Staubli VAL3: getTrajList.pgx

public program getTrajList(string& x_sItem[], num x_nIndex)
  local trsf l_tTrsf
  local string l_sItem[6]
  local string l_sEvent
  local string l_sItem2[7]
  local string l_sKey
  local num i
begin
  //  //获取列表
  //  resize(x_sItem,1,1)
  //  l_sKey=first(pt:tCommonStruct)
  //  i=0
  //  while l_sKey!=""
  //    if i!=0
  //      insert(x_sItem[i])
  //    endIf
  //    x_sItem[i]=l_sKey
  //    l_sKey=next(pt:tCommonStruct[l_sKey])
  //    i=i+1
  //    delay(0)
  //  endWhile
  //  if l_sKey=="" and i==0
  //    x_sItem[i]=""
  //  endIf

  //获取列表
  resize(x_sItem,1,x_nIndex)
  l_sKey=first(trajTemp:tTrajItem)
  i=0
  while l_sKey!=""
    x_sItem[i]=l_sKey
    l_sKey=next(trajTemp:tTrajItem[l_sKey])
    i=i+1
  endWhile
  if l_sKey=="" and i==0
    x_sItem[i]=""
  endIf
end
